(* IEC 61131-3 sources: brOscatLib/oscatBasic (part 7) *)

(* ---- STORE_8.st ---- *)
FUNCTION_BLOCK STORE_8
    (*http://www.oscat.de/images/OSCATBasic/oscat_basic333_en.pdf#page=253*)
    IF RST OR SET THEN
    	Q0 := NOT RST;
    	Q1 := Q0;
    	Q2 := Q0;
    	Q3 := Q0;
    	Q4 := Q0;
    	Q5 := Q0;
    	Q6 := Q0;
    	Q7 := Q0;
    ELSE
    	IF D0 THEN Q0 := TRUE; END_IF
    	IF D1 THEN Q1 := TRUE; END_IF
    	IF D2 THEN Q2 := TRUE; END_IF
    	IF D3 THEN Q3 := TRUE; END_IF
    	IF D4 THEN Q4 := TRUE; END_IF
    	IF D5 THEN Q5 := TRUE; END_IF
    	IF D6 THEN Q6 := TRUE; END_IF
    	IF D7 THEN Q7 := TRUE; END_IF

    	IF CLR AND NOT edge_ THEN
    		IF Q0 THEN Q0 := FALSE;
    		ELSIF Q1 THEN Q1 := FALSE;
    		ELSIF Q2 THEN Q2 := FALSE;
    		ELSIF Q3 THEN Q3 := FALSE;
    		ELSIF Q4 THEN Q4 := FALSE;
    		ELSIF Q5 THEN Q5 := FALSE;
    		ELSIF Q6 THEN Q6 := FALSE;
    		ELSE Q7 := FALSE;
    		END_IF
    	END_IF
    	edge_ := CLR;
    END_IF

    (* revision history
    hm	25.12.2007	rev 1.0
    	original version

    hm	30. oct. 2008	rev 1.1
    	optimized performance

    hm	14. mar. 2009	rev 1.2
    	removed double assignments

    *)

END_FUNCTION_BLOCK

(* ---- SUN_POS.st ---- *)
FUNCTION_BLOCK SUN_POS
    (*http://www.oscat.de/images/OSCATBasic/oscat_basic333_en.pdf#page=138*)

    (* n is the julian date and the number of days since 1.1.2000-12:00 midday *)
    (* be careful for step7 date startes 1.1.1990 instead of 1.1.1970 *)
    (* for step7 this line must change *)
    n := UDINT_TO_REAL(DT_TO_UDINT(UTC) - 946728000) * 0.000011574074074074;
    g :=MODR(6.240040768 + 0.01720197 * n, cPI2);
    d := MODR(4.89495042 + 0.017202792 * n, cPI2) + 0.033423055 * SIN(g) + 0.000349066 * SIN(2.0*g);
    e := 0.409087723 - 0.000000006981317008 * n;
    cos_d := COS(d);
    sin_d := SIN(d);
    a := ATAN(COS(e) * sin_d / cos_d);
    IF cos_d < 0.0 THEN a := a + cPI; END_IF
    c := ASIN(SIN(e) * sin_d);

    (* also here we must be very careful UTC is from 1.1.1970 for step7 the formula must change *)
    tau := RAD(MODR(6.697376 + (n - 0.25) * 0.0657098245037645 + UDINT_TO_REAL(TOD_TO_UDINT(DT_TO_TOD(UTC))) * 0.0000002785383333, 24.0) * 15.0 + LONGITUDE) - a;
    rlat := RAD(LATITUDE);
    sin_lat := SIN(rlat);
    cos_lat := COS(rlat);
    cos_tau := COS(tau);
    t1 := cos_tau * sin_lat - TAN(c) * cos_lat;
    B := ATAN(SIN(tau) / t1);
    IF t1< 0.0 THEN B := B + cPI2; ELSE B := B + cPI; END_IF
    B := DEG(MODR(B, cPI2));
    H := DEG(ASIN(COS(c) * cos_tau * cos_lat +SIN(c) * sin_lat));
    IF H > 180.0 THEN H := H - 360.0; END_IF
    (* consider refraction *)
    HR := H + REFRACTION(H);

    (* revision history
    hm	1. feb 2007	rev 1.0
    	original version

    hm	6. jan 2008	rev 1.1
    	performance improvements

    hm	18. jan 2008	rev 1.2
    	further performance improvements
    	only calculate once every 10 seconds

    hm	16. mar. 2008	rev 1.3
    	added type conversion to avoid warnings under codesys 3.0

    hm	30. jun. 2008	rev 1.4
    	added type conversions to avoid warnings under codesys 3.0

    hm	18. oct. 2008	rev 1.5
    	using math constants

    hm	17. dec. 2008	rev 1.6
    	angles below horizon are displayed in negative degrees

    hm	27. feb. 2009	rev 2.0
    	new code with better accuracy

    hm	7. mar. 2009	rev 2.1
    	refraction is added after angle normalization
    	deleted 10 second lockout
    	added output for astronomical heigth H
    *)
END_FUNCTION_BLOCK

(* ---- SUN_TIME.st ---- *)
FUNCTION_BLOCK SUN_TIME
    (*http://www.oscat.de/images/OSCATBasic/oscat_basic333_en.pdf#page=139*)
    b := LATITUDE * 0.0174532925199433;
    MIDDAY := SUN_MIDDAY(LONGITUDE, UTC);
    dk := 0.40954 * SIN(0.0172 * (INT_TO_REAL(DAY_OF_YEAR(UTC)) - 79.35));
    SUN_DECLINATION := DEG(dk);
    IF SUN_DECLINATION > 180.0 THEN SUN_DECLINATION := SUN_DECLINATION - 360.0; END_IF
    SUN_DECLINATION := 90.0 - LATITUDE + SUN_DECLINATION;
    delta := HOUR_TO_TIME(ACOS((SIN(RAD(H)) - SIN(b) * SIN(dk)) / (COS(b) * COS(dk))) * 3.819718632);
    SUN_RISE := MIDDAY - delta;
    SUN_SET := MIDDAY + delta;

    (* revision history

    rev 1.1	hm	20.1.2007
    	deleted unused variables sun_riseR and sun_setR

    rev 1.2 hm 17.4.2007
    	corrected error while sun:MIDDAY would not be corrected for LONGITUDE.

    rev 1.3	hm	6. jan 2008
    	performance improvements

    rev	1.4 hm	17. jan 2008
    	calculation is now only performed once a day

    hm	10. mar. 2009	rev 1.5
    	improved performance
    	calculation will be performed on every call to allow movong installations

    hm	26. jul 2009	rev 1.6
    	fixed a problem with wrong MIDDAY calculation

    hm	25. jan. 2011	rev 1.7
    	using function sun_midday
    	corrected angle of SUN_DECLINATION
    	added input H
    *)
END_FUNCTION_BLOCK

(* ---- TC_MS.st ---- *)
FUNCTION_BLOCK TC_MS
    (*http://www.oscat.de/images/OSCATBasic/oscat_basic333_en.pdf#page=352*)
    (* read system timer *)
    tx := T_PLC_MS();

    IF NOT init THEN
    	init := TRUE;
    	TC := 0;
    ELSE
    	TC := tx - last;
    END_IF
    last := tx;

    (* revision history
    hm		13. mar. 2008	rev 1.0
    	original version

    *)

END_FUNCTION_BLOCK

(* ---- TC_S.st ---- *)
FUNCTION_BLOCK TC_S
    (*http://www.oscat.de/images/OSCATBasic/oscat_basic333_en.pdf#page=353*)
    (* read system timer *)
    tx := T_PLC_US();

    IF NOT init THEN
    	init := TRUE;
    	TC := 0.0;
    ELSE
    	TC := UDINT_TO_REAL(tx - last)*1.0E-6;
    END_IF
    last := tx;

    (* revision history
    hm	13. mar. 2008	rev 1.0
    	original version

    hm	16. mar 2008	rev 1.1
    	added type conversion to avoid warnings under codesys 3.0

    hm	11. mar. 2009	rev 1.2
    	changed real constants to use dot syntax

    *)

END_FUNCTION_BLOCK

(* ---- TC_US.st ---- *)
FUNCTION_BLOCK TC_US
    (*http://www.oscat.de/images/OSCATBasic/oscat_basic333_en.pdf#page=353*)
    (* read system timer *)
    tx := T_PLC_US();

    IF NOT init THEN
    	init := TRUE;
    	TC := 0;
    ELSE
    	TC := tx - last;
    END_IF
    last := tx;

    (* revision history
    hm		13. mar. 2008	rev 1.0
    	original version

    *)

END_FUNCTION_BLOCK

(* ---- TEMPERATURE.st ---- *)
FUNCTION_BLOCK TEMPERATURE
    (*http://www.oscat.de/images/OSCATBasic/oscat_basic333_en.pdf#page=374*)
    YK := K + (C + 273.15) + (F + 459.67) * 0.555555555555 + (RE * 1.25 + 273.15) + (RA * 0.555555555555);
    YC := YK -273.15;
    YF := YK * 1.8 - 459.67;
    YRE := (YK - 273.15) * 0.8;
    YRA := YK * 1.8;

    (* revision history
    hm	21. feb. 2008	rev 1.0
    	original version

    *)
END_FUNCTION_BLOCK

(* ---- TICKER.st ---- *)
FUNCTION_BLOCK TICKER
    (*http://www.oscat.de/images/OSCATBasic/oscat_basic333_en.pdf#page=178*)

    (* generate next ticker when delay is low *)
    IF N < LEN(TEXT) THEN
    	IF NOT delay.Q THEN
    		(* increase step for next tick *)
    		step := step + 1;
    		IF step > LEN(TEXT) THEN step := 1; END_IF
    		(* extract dispay from TEXT *)
    		DISPLAY := MID(TEXT, N, step);
    		(* set delay timer for next tick *)
    		delay(IN := TRUE, PT := PT);
    	ELSE;
    		(* execute delay timer *)
    		delay(IN := FALSE);
    	END_IF
    ELSE
    	DISPLAY := TEXT;
    END_IF
    (* revision history
    hm	4. dec. 2007	rev 1.0
    	original version

    hm	15. dec. 2007	rev 1.1
    	step now starts at 1 instaed of 0

    hm	29. mar. 2008	rev 1.2
    	changed STRING to STRING(STRING_LENGTH)
    *)
END_FUNCTION_BLOCK

(* ---- TMAX.st ---- *)
FUNCTION_BLOCK TMAX
    (*http://www.oscat.de/images/OSCATBasic/oscat_basic333_en.pdf#page=204*)
    (* read system timer *)
    tx := UDINT_TO_TIME(T_PLC_MS());

    Z := FALSE;

    IF NOT IN THEN
    	Q := FALSE;
    ELSIF IN AND NOT last_in THEN
    	Q := TRUE;
    	start := tx;
    ELSIF (tx - start >= PT) AND Q THEN
    	Q := FALSE;
    	Z := TRUE;
    END_IF

    last_in := IN;

    (* revision history
    hm	20. jul. 2008	rev 1.0
    	original version

    *)
END_FUNCTION_BLOCK

(* ---- TMIN.st ---- *)
FUNCTION_BLOCK TMIN
    (*http://www.oscat.de/images/OSCATBasic/oscat_basic333_en.pdf#page=205*)
    pm(IN := IN, PT := PT);
    Q := IN OR pm.Q;

    (* revision history
    hm	21. jul. 2008	rev 1.0
    	original version

    *)
END_FUNCTION_BLOCK

(* ---- TOF_1.st ---- *)
FUNCTION_BLOCK TOF_1
    (*http://www.oscat.de/images/OSCATBasic/oscat_basic333_en.pdf#page=205*)
    (* read system timer *)
    tx := UDINT_TO_TIME(T_PLC_MS());

    IF RST THEN
    	Q := FALSE;
    ELSIF IN THEN
    	Q := TRUE;
    	start := tx;
    ELSIF tx - start >= PT THEN
    	Q := FALSE;
    END_IF

    (* revision history
    hm	17. jul. 2008	rev 1.0
    	original version

    *)
END_FUNCTION_BLOCK

(* ---- TOGGLE.st ---- *)
FUNCTION_BLOCK TOGGLE
    (*http://www.oscat.de/images/OSCATBasic/oscat_basic333_en.pdf#page=254*)
    IF RST THEN
    	Q := 0;
    ELSIF CLK AND NOT edge_ THEN
    	Q := NOT Q;
    END_IF
    edge_ := CLK;

    (* revision history

    hm	13.9.2007		rev 1.0
    	original version

    hm	30. oct. 2008	rev 1.1
    	deleted unnecessary init

    *)

END_FUNCTION_BLOCK

(* ---- TONOF.st ---- *)
FUNCTION_BLOCK TONOF
    (*http://www.oscat.de/images/OSCATBasic/oscat_basic333_en.pdf#page=206*)
    IF IN XOR old THEN
      X(IN := FALSE, PT := SEL(IN,T_OFF,T_ON));
      mode := IN;
      old := IN;
    END_IF
    X(IN := TRUE);
    IF X.Q THEN Q := mode;END_IF

    (* revision history
    hm	10. dec 2007	rev 1.0
    	original version

    hm	17. sep. 2007	rev 1.1
    	improved performance

    hm	21. jul. 2009	rev 1.2
    	fixed a timing probelm

    *)

END_FUNCTION_BLOCK

(* ---- TP_1.st ---- *)
FUNCTION_BLOCK TP_1
    (*http://www.oscat.de/images/OSCATBasic/oscat_basic333_en.pdf#page=207*)
    (* read system timer *)
    tx := UDINT_TO_TIME(T_PLC_MS());

    IF RST THEN
    	Q := FALSE;
    ELSIF IN AND NOT ix THEN
    	Q := TRUE;
    	start := tx;
    ELSIF tx - start >= PT THEN
    	Q := FALSE;
    END_IF

    ix:= IN;

    (* revision history
    hm	28. jun. 2008
    	original version

    *)
END_FUNCTION_BLOCK

(* ---- TP_1D.st ---- *)
FUNCTION_BLOCK TP_1D
    (*http://www.oscat.de/images/OSCATBasic/oscat_basic333_en.pdf#page=208*)
    (* read system timer *)
    tx := UDINT_TO_TIME(T_PLC_MS());

    IF RST THEN
    	Q := FALSE;
    	RST := FALSE;
    	W := FALSE;
    ELSIF W THEN
    	IF tx - start >= PTD THEN
    		W := FALSE;
    	END_IF
    ELSIF IN AND NOT ix THEN
    	Q := TRUE;
    	start := tx;
    	IN := FALSE;
    ELSIF tx - start >= PT1 THEN
    	Q := FALSE;
    	W := TRUE;
    	start := tx;
    END_IF

    ix := IN;

    (* revision history
    hm	28. jun. 2008
    	original version

    *)
END_FUNCTION_BLOCK

(* ---- TP_X.st ---- *)
FUNCTION_BLOCK TP_X
    (*http://www.oscat.de/images/OSCATBasic/oscat_basic333_en.pdf#page=208*)
    (* read system_time *)
    tx := UDINT_TO_TIME(T_PLC_MS());

    (* rising edge_ trigger *)
    IF IN AND NOT edge_ THEN
    	start := tx;
    	Q := PT > t#0ms;
    ELSIF Q THEN
    	ET := tx - start;
    	IF ET >= PT THEN
    		Q := FALSE;
    		ET := t#0ms;
    	END_IF
    END_IF
    edge_ := IN;

    (* revision history
    hm	4. aug 2006		rev 1.0
    	original version

    hm	17. sep 2007	rev 1.1
    	replaced time() with T_PLC_MS() for compatibility reasons

    hm	19. oct. 2008	rev 1.2
    	renamed to TP_R to TP_X for compatibility reasons

    hm	17. dec. 2008	rev 1.3
    	code optimized

    *)
END_FUNCTION_BLOCK

(* ---- TREND.st ---- *)
FUNCTION_BLOCK TREND
    (*http://www.oscat.de/images/OSCATBasic/oscat_basic333_en.pdf#page=305*)
    TU := X > last_X;
    TD := X < last_X;
    Q := TU OR TD;
    D := X - last_X;

    last_X := X;

    (* revision history
    hm	21. aug. 2009	rev 1.0
    	original version

    *)

END_FUNCTION_BLOCK

(* ---- TREND_DW.st ---- *)
FUNCTION_BLOCK TREND_DW
    (*http://www.oscat.de/images/OSCATBasic/oscat_basic333_en.pdf#page=315*)
    IF DWORD_TO_UDINT(X) > last_X THEN
    	TU := TRUE;
    	TD := FALSE;
    	D := UDINT_TO_DWORD(DWORD_TO_UDINT(X) - last_X);
    	Q := TRUE;
    ELSIF DWORD_TO_UDINT(X) < last_X THEN
    	TD := TRUE;
    	TU := FALSE;
    	D := UDINT_TO_DWORD(last_X - DWORD_TO_UDINT(X));
    	Q := FALSE;
    ELSE
    	TU := FALSE;
    	TD := FALSE;
    	D := 0;
    END_IF
    last_X := DWORD_TO_UDINT(X);

    (* revision history
    hm	21. nov. 2008	rev 1.0
    	original version

    hm	20. feb. 2009	rev 1.1
    	added outputs TU, TD and D

    hm	14. mar. 2009	rev 1.2
    	removed double assignments

    *)

END_FUNCTION_BLOCK

(* ---- TUNE.st ---- *)
FUNCTION_BLOCK TUNE
    (*http://www.oscat.de/images/OSCATBasic/oscat_basic333_en.pdf#page=472*)
    (* read system time *)
    tx := T_PLC_MS();

    IF RST THEN
    	Y := RST_VAL;
    	state := 0;
    ELSIF SET THEN
    	Y := SET_VAL;
    	state := 0;
    ELSIF state > 0 THEN
    	(* key has been pushed state machine operating *)
    	(* first read the correct input *)
    	IF state = 1 THEN
    		(* step up *)
    		in := SU;
    	ELSE
    		(* step down *)
    		in := SD;
    	END_IF
    	(* check for single step operation *)
    	IF NOT in AND tx - start <= TIME_TO_UDINT(T1) THEN
    		Y := Y_start + step;
    		state := 0;
    	(* check if fast ramp needs to be generated *)
    	ELSIF in AND tx - start >= TIME_TO_UDINT(T2) THEN
    		Y := Y_start2 + UDINT_TO_REAL(tx - start2) * S2 / SPEED;
    	(* check if slow ramp needs to be generated *)
    	ELSIF in AND tx - start >= TIME_TO_UDINT(T1) THEN
    		Y := Y_start + UDINT_TO_REAL(tx - start - TIME_TO_UDINT(T1)) * S1 / SPEED;
    		start2 := tx;
    		Y_start2 := Y;
    	ELSIF NOT in THEN
    		state := 0;
    	END_IF
    ELSIF SU THEN
    	(* slow step up *)
    	state := 1;
    	start := tx;
    	step := SS;
    	SPEED := 1000.0;
    	Y_start := Y;
    ELSIF SD THEN
    	(* slow step down *)
    	state := 2;
    	start := tx;
    	step := -SS;
    	SPEED := -1000.0;
    	Y_start := Y;
    END_IF

    (* make sure output does not exceed limits *)
    Y := LIMIT(LIMIT_L, Y, LIMIT_H);

    (* revision history
    hm	3.11.2007		rev 1.0
    	original version

    hm	16. mar. 2008	rev 1.1
    	added type conversions to avoid warnings under codesys 3.0

    hm	11. mar. 2009	rev 1.2
    	real constants updated to new systax using dot

    *)
END_FUNCTION_BLOCK

(* ---- TUNE2.st ---- *)
FUNCTION_BLOCK TUNE2
    (*http://www.oscat.de/images/OSCATBasic/oscat_basic333_en.pdf#page=475*)
    (* read system time *)
    tx := T_PLC_MS();

    IF RST THEN
    	Y := RST_VAL;
    	state := 0;
    ELSIF SET THEN
    	Y := SET_VAL;
    	state := 0;
    ELSIF state > 0 THEN
    	(* key has been pushed state machine operating *)
    	(* first read the correct input *)
    	CASE state OF
    		1 :	(* slow up *)
    			in := SU;
    		2 :	(* slow down *)
    			in := SD;
    		3 :	(* fast up *)
    			in := FU;
    		4 :	(* fast down *)
    			in := FD;
    	END_CASE
    	(* check for single step operation *)
    	IF NOT in AND tx - start <= TIME_TO_UDINT(TR) THEN
    		Y := Y_start + step;
    		state := 0;
    	(* check if ramp needs to be generated *)
    	ELSIF in AND tx - start >= TIME_TO_UDINT(TR) THEN
    		Y := Y_start + UDINT_TO_REAL(tx - start - TIME_TO_UDINT(TR)) * SPEED;
    	ELSIF NOT in THEN
    		state := 0;
    	END_IF
    ELSIF SU THEN
    	(* slow step up *)
    	state := 1;
    	start := tx;
    	step := SS;
    	SPEED := S1 * 1.0E-3;
    	Y_start := Y;
    ELSIF SD THEN
    	(* slow step down *)
    	state := 2;
    	start := tx;
    	step := -SS;
    	SPEED := -S1 * 1.0E-3;
    	Y_start := Y;
    ELSIF FU THEN
    	(* fast step up *)
    	state := 3;
    	start := tx;
    	step := FS;
    	SPEED := S2 * 1.0E-3;
    	Y_start := Y;
    ELSIF FD THEN
    	(* fast step down *)
    	state := 4;
    	start := tx;
    	step := -FS;
    	SPEED := -S2 * 1.0E-3;
    	Y_start := Y;
    END_IF

    (* make sure output does not exceed limits *)
    Y := LIMIT(LIMIT_L, Y, LIMIT_H);

    (* revision history
    hm	3.11.2007		rev 1.0
    	original version

    hm	16. 3. 2008	rev 1.1
    	added type conversions to avoid warnings in codesys 3.0
    	improved performance

    hm	11. mar. 2009	rev 1.2
    	real constants updated to new systax using dot

    *)
END_FUNCTION_BLOCK

(* ---- oscatBasic.var ---- *)
VAR CONSTANT
	STRING_LENGTH : INT := 250;
	cCHARNAMES : ARRAY[1..4] OF STRING[253] := [';"&quot;&&amp;<&lt;>&gt;€&euro; &nbsp;¡&iexcl;¢&cent;£&pound;¤&curren;¥&yen;¦&brvbar;§&sect;¨&uml;©&copy;ª&ordf;«&laquo;¬&not;­&shy;®&reg;¯&macr;°&deg;±&plusmn;²&sup2;³&sup3;´&acute;µ&micro;¶&para;·&middot;¸&cedil;¹&sup1;º&ordm;»&raquo;¼&frac14;Û&Ucirc;',
		';¾&frac34;¿&iquest;À&Agrave;Á&Aacute;Â&Acirc;Ã&Atilde;Ä&Auml;Å&Aring;Æ&AElig;Ç&Ccedil;È&Egrave;É&Eacute;Ê&Ecirc;Ë&Euml;Ì&Igrave;Í&Iacute;Î&Icirc;Ï&Iuml;Ð&ETH;Ñ&Ntilde;Ò&Ograve;Ó&Oacute;Ô&Ocirc;Õ&Otilde;Ö&Ouml;×&times;Ø&Oslash;Ù&Ugrave;Ú&Uacute;½&frac12;',
		';Ü&Uuml;Ý&Yacute;Þ&THORN;ß&szlig;à&agrave;á&aacute;â&acirc;ã&atilde;ä&auml;å&aring;æ&aelig;ç&ccedil;è&egrave;é&eacute;ê&ecirc;ë&euml;ì&igrave;í&iacute;î&icirc;ï&iuml;ð&eth;ñ&ntilde;ò&ograve;ó&oacute;ô&ocirc;õ&otilde;ö&ouml;÷&divide;ø&oslash;ù&ugrave;',
		';ú&uacute;û&ucirc;ü&uuml;ý&yacute;þ&thorn;ÿ&yuml;'];
	cMTH_OFS : ARRAY[1..12] OF INT := [0,31,59,90,120,151,181,212,243,273,304,334]; (*Setup - Month offsets*)
	cDECADES : ARRAY[0..8] OF REAL := [1,10,100,1000,10000,100000,1000000,10000000,100000000]; (*Setup - Decades*)
	cLOCATION_DEFAULT : INT := 1; (* Location - 1=germany, 2=austria 3=france 4=belgium-german 5= italien-Südtirol *)
	cLOCATION_LMAX : INT := 5; (* Location - ?? *)
	cLOCATION_LANGUAGE : ARRAY[1..5] OF INT := [2,2,3,2,2]; (* Location - language spoken in the location *)
	cEXTENDED_ASCII : BOOL := TRUE; (*Setup - Extended ascii enabled*)
	cLANGUAGE_DEFAULT : INT := 1; (* 1=english, 2=german 3=french *)
	cLANGUAGE_WEEKDAYS : ARRAY[1..3,1..7] OF STRING[10] := ['Monday','Tuesday','Wednesday','Thursday','Friday','Saturday','Sunday','Montag','Dienstag','Mittwoch','Donnerstag','Freitag','Samstag','Sonntag','Lundi','Mardi','Mercredi','Jeudi','Vendredi','Samedi','Dimanche'];
	cLANGUAGE_WEEKDAYS2 : ARRAY[1..3,1..7] OF STRING[2] := ['Mo','Tu','We','Th','Fr','Sa','Su','Mo','Di','Mi','Do','Fr','Sa','So','Lu','Ma','Me','Je','Ve','Sa','Di'];
	cLANGUAGE_MONTHS : ARRAY[1..3,1..12] OF STRING[10] := ['January','February','March','April','May','June','July','August','September','October','November','December','Januar','Februar','März','April','Mai','Juni','Juli','August','September','Oktober','November','Dezember','Janvier','Février','mars','Avril','Mai','Juin','Juillet','Août','Septembre','Octobre','Novembre','Decembre'];
	cLANGUAGE_MONTHS3 : ARRAY[1..3,1..12] OF STRING[3] := ['Jan','Feb','Mar','Apr','May','Jun','Jul','Aug','Sep','Oct','Nov','Dec','Jan','Feb','Mrz','Apr','Mai','Jun','Jul','Aug','Sep','Okt','Nov','Dez','Jan','Fev','Mar','Avr','Mai','Jun','Jul','Aou','Sep','Oct','Nov','Dec'];
	cLANGUAGE_DIRS : ARRAY[1..3,0..15] OF STRING[3] := ['N','NNE','NE','ENE','E','ESE','SE','SSE','S','SSW','SW','WSW','W','WNW','NW','NNW','N','NNO','NO','ONO','O','OSO','SO','SSO','S','SSW','SW','WSW','W','WNW','NW','NNW','N','NNO','NO','ONO','O','OSO','SO','SSO','S','SSW','SW','WSW','W','WNW','NW','NNW'];
	LANGUAGE : CONSTANTS_LANGUAGE := (DEFAULT:=1,LMAX:=3,WEEKDAYS:=['Monday','Tuesday','Wednesday','Thursday','Friday','Saturday','Sunday','Montag','Dienstag','Mittwoch','Donnerstag','Freitag','Samstag','Sonntag','Lundi','Mardi','Mercredi','Jeudi','Vendredi','Samedi','Dimanche'],WEEKDAYS2:=['Mo','Tu','We','Th','Fr','Sa','Su','Mo','Di','Mi','Do','Fr','Sa','So','Lu','Ma','Me','Je','Ve','Sa','Di'],MONTHS:=['January','February','March','April','May','June','July','August','September','October','November','December','Januar','Februar','MÃƒÂ¤rz','April','Mai','Juni','Juli','August','September','Oktober','November','Dezember','Janvier','FÃƒÂ©vrier','mars','Avril','Mai','Juin','Juillet','AoÃƒÂ»t','Septembre','Octobre','Novembre','Decembre'],MONTHS3:=['Jan','Feb','Mar','Apr','May','Jun','Jul','Aug','Sep','Oct','Nov','Dec','Jan','Feb','Mrz','Apr','Mai','Jun','Jul','Aug','Sep','Okt','Nov','Dez','Jan','Fev','Mar','Avr','Mai','Jun','Jul','Aou','Sep','Oct','Nov','Dec'],DIRS:=['N','NNE','NE','ENE','E','ESE','SE','SSE','S','SSW','SW','WSW','W','WNW','NW','NNW','N','NNO','NO','ONO','O','OSO','SO','SSO','S','SSW','SW','WSW','W','WNW','NW','NNW','N','NNO','NO','ONO','O','OSO','SO','SSO','S','SSW','SW','WSW','W','WNW','NW','NNW']); (*Language constants*)
	cLANGUAGE_LMAX : INT := 3;
	cPN : REAL := 8.314472; (*Physics constants - Atmospheric pressure*)
	cR : REAL := 8.314472; (*Physics constants - Gas constant*)
	cT0 : REAL := -273.15; (*Physics constants - Celsius at 0K*)
	LIST_LENGTH : INT := 250;
	MATH : CONSTANTS_MATH := (PI:=3.1415926535897931,PI2:=6.2831853071795862,PI4:=12.566370614359172,PI05:=1.5707963267949,PI025:=0.785398163397448,PI_INV:=0.318309886183791,E:=2.7182818284590451,E_INV:=0.367879441171442,SQ2:=1.4142135623731,FACTS:=[1,1,2,6,24,120,720,5040,40320,362880,3628800,39916800,479001600]); (*Math constants*)
	cPI : REAL := 3.1415926535897931; (*Math constants - PI*)
	cPI2 : REAL := 6.2831853071795862; (*Math constants - PI*2*)
	cPI4 : REAL := 12.566370614359172; (*Math constants - PI*4*)
	cPI05 : REAL := 1.5707963267949; (*Math constants - PI / 2*)
	cPI025 : REAL := 0.785398163397448; (*Math constants - PI / 4*)
	cPI_INV : REAL := 0.318309886183791; (*Math constants - Inverse PI number*)
	ce : REAL := 2.7182818284590451; (*Math constants - Eulers number*)
	ce_INV : REAL := 0.367879441171442; (*Math constants - Inverse eulers number*)
	cSQ2 : REAL := 1.4142135623731; (*Math constants - Square root of 2*)
	PHYS : CONSTANTS_PHYS := (C:=299792458,E:=1.60217653E-19,G:=9.80665,T0:=-273.15,RU:=8.314472,PN:=101325); (*Physics constants*)
	cC : REAL := 299792458; (*Physics constants - Speed of light*)
	cE : REAL := 1.60217653E-19; (*Physics constants - Mass energy*)
	cg : REAL := 9.80665; (*Physics constants - Gravitational acceleration on Earth*)
	SETUP : CONSTANTS_SETUP := (EXTENDED_ASCII:=TRUE,CHARNAMES:=['1'],MTH_OFS:=[0,31,59,90,120,151,181,212,243,273,304,334]); (*Setup constants*)
	LOCATION : CONSTANTS_LOCATION := (DEFAULT:=1,LMAX:=5,LANGUAGE:=[2(2),3,2(2)]); (*Location constants*)
END_VAR
